Fanuc KAREL source: KO00026.KL

PROGRAM KO00026
%NOLOCKGROUP
VAR
  P1: JOINTPOS
  P2: JOINTPOS
  P3: JOINTPOS
  OUT: XYZWPR
BEGIN
  OUT = FRAME(P1, P2, P3)
END KO00026
